(* PLC project g_batch_mixer_clean, Anonymous Benchmark Suite 1.0 *)
(* stored: creationDateTime 2026-07-09T00:00:00 *)

PROGRAM g_batch_mixer_clean
  VAR_INPUT
    mix_cmd : BOOL;
    lid_open : BOOL;
    enable : BOOL;
    maint : BOOL;
  END_VAR
  VAR_OUTPUT
    mixer : BOOL;
    alarm : BOOL;
  END_VAR

(* LD diagram, written out as Structured Text *)
mixer := NOT lid_open AND mix_cmd AND enable;
alarm := lid_open;
END_PROGRAM

CONFIGURATION Config0
  RESOURCE Res0 ON PLC
    TASK tcyclic(INTERVAL := T#10ms, PRIORITY := 0);
    PROGRAM inst0 WITH tcyclic : g_batch_mixer_clean;
  END_RESOURCE
END_CONFIGURATION
